// TIA Portal V21 export
// export: Created 2026-11-22T02:34:23.7994351Z, ExportSetting WithDefaults, DisplayName Totally Integrated Automation Portal, DisplayVersion V21 Update 3, DisplayName STEP 7 Professional, DisplayVersion V21 Update 3, DisplayName STEP 7 Safety, DisplayVersion V21, DisplayName Tech WebApplication, DisplayVersion V21, DisplayName WinCC Basic/Comfort/Advanced, DisplayVersion V21 Update 3, DisplayName WinCC Unified, DisplayVersion V21 Update 3
VBScript "SetS2"  Type=Sub
  SmartTags("D_State") = 2
  SmartTags("D_Bool") = True
  SmartTags("D_SInt") = 12
  SmartTags("D_Int") = 1234
  SmartTags("D_DInt") = 123456
  SmartTags("D_USInt") = 200
  SmartTags("D_UInt") = 40000
  SmartTags("D_UDInt") = 3000000000
  SmartTags("D_Real") = 3.14159
  SmartTags("D_LReal") = 2.718281828
  SmartTags("D_String") = "Hello World"
  SmartTags("D_DateTime") = DateSerial(2026, 11, 22) + TimeSerial(13, 45, 30)
  SmartTags("D_Pct") = 50
  SmartTags("D_Range") = 25
  SmartTags("D_Bits") = 2
  SmartTags("D_Vis") = True
  SmartTags("D_En") = True
  SmartTags("D_X") = 200
  SmartTags("D_Y") = 120
  SmartTags("D_Max") = 200
  SmartTags("D_Min") = -100
  SmartTags("D_TL") = 5
  SmartTags("D_BarR") = 0
